Universal Robots URScript: SpeedProg.script

def SpeedProg():
  # Global parameters:
  global speed_ms    = 0.250
  global speed_rads  = 0.750
  global accel_mss   = 1.200
  global accel_radss = 1.200
  global blend_radius_m = 0.001
  global ref_frame = p[0,0,0,0,0,0]

  #
  # TO REMOVE HEADER:
  # Go to "Program" -> "Post-Processor Editor"
  # Select "Universal Robots"
  # Set "INCLUDE_HEADER" to "False"
  #
  #--------------------------
  # Add any default subprograms here
  # For example, to drive a gripper as a program call:
  # def Gripper_Open():
  #   ...
  # end
  #
  # Example to drive a spray gun:
  def SprayOn(value):
    # use the value as an output:
    DO_SPRAY = 5
    if value == 0:
      set_standard_digital_out(DO_SPRAY, False)
    else:
      set_standard_digital_out(DO_SPRAY, True)
    end
  end

  # Example to drive an extruder:
  def Extruder(value):
    # use the value as an output:
    if value < 0:
      # stop extruder
    else:
      # start extruder
    end
  end

  # Example to move an external axis
  def MoveAxis(value):
    # use the value as an output:
    DO_AXIS_1 = 1
    DI_AXIS_1 = 1
    if value <= 0:
      set_standard_digital_out(DO_AXIS_1, False)

      # Wait for digital input to change state
      #while (get_standard_digital_in(DI_AXIS_1) != False):
      #  sync()
      #end
    else:
      set_standard_digital_out(DO_AXIS_1, True)

      # Wait for digital input to change state
      #while (get_standard_digital_in(DI_AXIS_1) != True):
      #  sync()
      #end
    end
  end
  #--------------------------


  # Main program:
  # Program generated by RoboDK v6.0.7 for UR10 on XX/XX/XXXX 18:00:00
  # Using nominal kinematics.
  ref_frame = p[1.234570, -0.098765, 0.050500, 0.000000, 0.000000, 0.523599]
  set_tcp(p[0.010000, 0.020000, 0.150000, 0.000000, 0.000000, 0.000000])
  blend_radius_m = 0.000
  speed_ms    = 0.001
  movel(pose_trans(ref_frame,p[-0.607850, 0.543849, 0.363215, 0.731956, 2.185937, -0.570291]),accel_mss,speed_ms,t=0,r=0)
  speed_rads  = 0.017
  movej([0.000000, -0.174533, 0.349066, 0.000000, 0.523599, 0.000000],accel_radss,speed_rads,t=0,r=0)
  blend_radius_m = 0.001
  speed_ms    = 0.012
  movel(pose_trans(ref_frame,p[-0.640584, 0.506980, 0.371534, 0.731956, 2.185937, -0.570291]),accel_mss,speed_ms,t=0,r=0)
  speed_rads  = 0.096
  movej([0.349066, -0.174533, 0.349066, 0.000000, 0.523599, 0.000000],accel_radss,speed_rads,t=0,r=0)
  blend_radius_m = 0.003
  speed_ms    = 0.100
  movel(pose_trans(ref_frame,p[-0.607850, 0.543849, 0.363215, 0.731956, 2.185937, -0.570291]),accel_mss,speed_ms,t=0,r=0)
  speed_rads  = 0.349
  movej([0.000000, -0.174533, 0.349066, 0.000000, 0.523599, 0.000000],accel_radss,speed_rads,t=0,r=0)
  blend_radius_m = 0.004
  speed_ms    = 0.333
  movel(pose_trans(ref_frame,p[-0.640584, 0.506980, 0.371534, 0.731956, 2.185937, -0.570291]),accel_mss,speed_ms,t=0,r=0)
  speed_rads  = 0.785
  movej([0.349066, -0.174533, 0.349066, 0.000000, 0.523599, 0.000000],accel_radss,speed_rads,t=0,r=0)
  blend_radius_m = 0.006
  speed_ms    = 1.000
  movel(pose_trans(ref_frame,p[-0.607850, 0.543849, 0.363215, 0.731956, 2.185937, -0.570291]),accel_mss,speed_ms,t=0,r=0)
  speed_rads  = 1.571
  movej([0.000000, -0.174533, 0.349066, 0.000000, 0.523599, 0.000000],accel_radss,speed_rads,t=0,r=0)
  blend_radius_m = 0.009
  speed_ms    = 2.500
  movel(pose_trans(ref_frame,p[-0.640584, 0.506980, 0.371534, 0.731956, 2.185937, -0.570291]),accel_mss,speed_ms,t=0,r=0)
  speed_rads  = 2.094
  movej([0.349066, -0.174533, 0.349066, 0.000000, 0.523599, 0.000000],accel_radss,speed_rads,t=0,r=0)
  blend_radius_m = 0.015
  speed_ms    = 3.000
  movel(pose_trans(ref_frame,p[-0.607850, 0.543849, 0.363215, 0.731956, 2.185937, -0.570291]),accel_mss,speed_ms,t=0,r=0)
  speed_rads  = 3.142
  movej([0.000000, -0.174533, 0.349066, 0.000000, 0.523599, 0.000000],accel_radss,speed_rads,t=0,r=0)
  blend_radius_m = 0.030
  movel(pose_trans(ref_frame,p[-0.640584, 0.506980, 0.371534, 0.731956, 2.185937, -0.570291]),accel_mss,speed_ms,t=0,r=0)
  speed_rads  = 3.142
  movej([0.349066, -0.174533, 0.349066, 0.000000, 0.523599, 0.000000],accel_radss,speed_rads,t=0,r=0)
  blend_radius_m = 0.075
  speed_ms    = 0.001
  movel(pose_trans(ref_frame,p[-0.607850, 0.543849, 0.363215, 0.731956, 2.185937, -0.570291]),accel_mss,speed_ms,t=0,r=0)
  speed_rads  = 3.142
  movej([0.000000, -0.174533, 0.349066, 0.000000, 0.523599, 0.000000],accel_radss,speed_rads,t=0,r=0)
  blend_radius_m = 0.150
  speed_ms    = 0.750
  movel(pose_trans(ref_frame,p[-0.640584, 0.506980, 0.371534, 0.731956, 2.185937, -0.570291]),accel_mss,speed_ms,t=0,r=0)
  speed_rads  = 0.039
  movej([0.349066, -0.174533, 0.349066, 0.000000, 0.523599, 0.000000],accel_radss,speed_rads,t=0,r=0)
  accel_mss   = 2.000
  accel_radss = 8.727
  movel(pose_trans(ref_frame,p[-0.640584, 0.506980, 0.371534, 0.731956, 2.185937, -0.570291]),accel_mss,speed_ms,t=0,r=0)
  # End of main program
end

SpeedProg()
